Universal Robots URScript: T008_codellama_34b_baseline_rep2_retry3.urscript

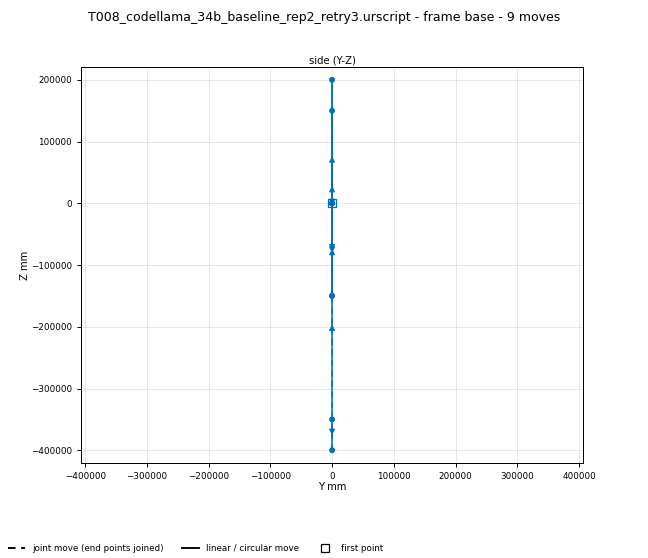
[picture p0: tool path of T008_codellama_34b_baseline_rep2_retry3.urscript in frame base, 9 of 9 moves have a stored position in this frame; points joined in program order, loops and branches not executed]
def heavy_depalletizing():
    # Home the robot arm
    movej(p[0, 0, 0, 0, 0, 0], v=400)

    # Move above the pallet
    movel(p[0, 0, 150, 0, 0, 0], v=400)

    # Descend to the top layer of the pallet
    movel(p[0, 0, -150, 0, 0, 0], v=150)

    # Lift the box off the pallet
    movel(p[0, 0, 200, 0, 0, 0], v=200)

    # Transit to the conveyor belt
    movel(p[0, 0, -350, 0, 0, 0], v=350)

    # Move along the conveyor belt
    movel(p[0, 0, -400, 0, 0, 0], v=400)

    # Place the box on the conveyor belt
    movej(p[0, 0, 0, 0, 0, 0], v=400)

    # Move back to the starting position
    movel(p[0, 0, -150, 0, 0, 0], v=200)

    # Lift the arm back up
    movej(p[0, 0, 0, 0, 0, 0], v=400)
